// TIA Portal V19 export
TYPE "ST_FENCE"
   STRUCT
      Safety_Fence_1 : Bool;
      Safety_Fence_2 : Bool;
      Safety_Fence_3 : Bool;
      Safety_Fence_4 : Bool;
      Safety_Fence_5 : Bool;
      Safety_Fence_6 : Bool;
      Safety_Fence_7 : Bool;
      Safety_Fence_8 : Bool;
      Safety_Fence_9 : Bool;
      Safety_Fence_10 : Bool;
   END_STRUCT;
END_TYPE
